(* IEC 61131-3 sources: Palletizer_Control_with_Automation_Studio/Task_1/Logical/Libraries/MpCom, 3 files *)

(* ---- MpCom.typ ---- *)
TYPE
	MpComConfigScopeEnum :
		(
		mpCOM_CONFIG_SCOPE_COMPONENT := 0, (*Import / Export configuration only for given component*)
		mpCOM_CONFIG_SCOPE_BRANCH := 1 (*Import / Export configuration for given component and all its sub-components*)
		);
	MpComStatusIDType : 	STRUCT
		ID : MpComErrorEnum; (*Status ID*)
		Severity : MpComSeveritiesEnum; (*Status severity*)
		Facility : MpComFacilitiesEnum; (*Status facility*)
		Code : UINT; (*Status / Error code*)
	END_STRUCT;
	MpComDiagType : 	STRUCT
		StatusID : MpComStatusIDType; (*StatusID diagnostic structure *)
	END_STRUCT;
	MpComConfigManagerInfoType : 	STRUCT
		Diag : MpComDiagType; (*Diagnostic structure for the status ID*)
	END_STRUCT;
	MpComDumpInternalType : 	STRUCT
		CmdOld : BOOL;
	END_STRUCT;
	MpComLoggerUISetupType : 	STRUCT
		LoggerListSize : UINT := 20; (*Number of logger entries to be displayed on one page of the list in the HMI application*)
		LoggerScrollWindow : USINT := 0; (*Determines how many entries from the list are displayed in advance when scrolling up and down*)
	END_STRUCT;
	MpComLoggerUIConnectType : 	STRUCT
		Status : MpComLoggerUIStatusEnum;
		List : MpComLoggerUILoggerListType; (*List of resultant logger entries*)
		Clear : BOOL; (*Clean the internal buffer*)
		SearchFilter : STRING[255]; (*Filter used to define the visibility of entries*)
	END_STRUCT;
	MpComLoggerUIStatusEnum :
		(
		mpCOM_LOGGERUI_IDLE := 0,
		mpCOM_LOGGERUI_REFRESH := 1,
		mpCOM_LOGGERUI_ERROR := 2
		);
	MpComLoggerUILoggerListType : 	STRUCT
		Message : ARRAY[0..19]OF STRING[255]; (*List of logger entries: message*)
		StatusID : ARRAY[0..19]OF DINT; (*List of logger entries: status ID*)
		ErrorNumber : ARRAY[0..19]OF UINT; (*List of logger entries: error code as part of Status ID*)
		Time : ARRAY[0..19]OF MpComLoggerUIDateTimeType; (*List of logger entries: date, time and microseconds*)
		Component : ARRAY[0..19]OF STRING[50]; (*List of logger entries: component name*)
		Facility : ARRAY[0..19]OF MpComFacilitiesEnum; (*List of logger entries: facility as part of Status ID*)
		Severity : ARRAY[0..19]OF MpComSeveritiesEnum; (*List of logger entries: severity as part of Status ID*)
		PageUp : BOOL; (*Jumps to the start of the current page and then scrolls up one page at a time *)
		PageDown : BOOL; (*Jumps to the end of the current page and then scrolls down one page at a time *)
		StepUp : BOOL; (*Selects the previous entry in the list*)
		StepDown : BOOL; (*Selects the next entry in the list*)
		RangeStart : REAL; (*Shows a bar indicating which part of the list is currently being displayed-Start [%]*)
		RangeEnd : REAL; (*Shows a bar indicating which part of the list is currently being displayed-End [%]*)
	END_STRUCT;
	MpComLoggerUIDateTimeType : 	STRUCT
		DateTime : DATE_AND_TIME; (*List of logger entries: date and time: the view could be customized on VC*)
		Microseconds : UDINT; (*List of logger entries: additional information about microseconds when the event was triggered*)
	END_STRUCT;
	MpComLoggerUIInfoType : 	STRUCT
		CurrentBufferEntries : UINT; (*Number of entries currently in the internal buffer. It is a ring buffer, it means that reached the BufferSize it doesn't increase any more*)
		Diag : MpComDiagType; (*Diagnostic structure for the status ID*)
	END_STRUCT;
END_TYPE

(* ---- MpComError.typ ---- *)
TYPE
    MpComErrorEnum :
        ( (* Error numbers of library MpCom *)
        mpCOM_NO_ERROR := 0, (* No error *)
        mpCOM_ERR_ACTIVATION := -1064239103, (* Could not create component [Error: 1, 0xc0910001] *)
        mpCOM_ERR_MPLINK_NULL := -1064239102, (* MpLink is NULL pointer [Error: 2, 0xc0910002] *)
        mpCOM_ERR_MPLINK_INVALID := -1064239101, (* MpLink connection not allowed [Error: 3, 0xc0910003] *)
        mpCOM_ERR_MPLINK_CHANGED := -1064239100, (* MpLink modified [Error: 4, 0xc0910004] *)
        mpCOM_ERR_MPLINK_CORRUPT := -1064239099, (* Invalid MpLink contents [Error: 5, 0xc0910005] *)
        mpCOM_ERR_LINK_NOT_POSSIBLE := -1064238848, (* Connection not possible [Error: 256, 0xc0910100] *)
        mpCOM_ERR_FILE_SYSTEM := -1064238847, (* Error editing file [Error: 257, 0xc0910101] *)
        mpCOM_ERR_INVALID_FILE_DEV := -1064238846, (* Invalid file device [Error: 258, 0xc0910102] *)
        mpCOM_ERR_INVALID_FILE_NAME := -1064238845, (* Invalid filename [Error: 259, 0xc0910103] *)
        mpCOM_ERR_NO_CONFIG_IMPORT := -1064238844, (* No configuration data was imported [Error: 260, 0xc0910104] *)
        mpCOM_ERR_MISSING_UICONNECT := -1064238843, (* Missing value on UIConnect [Error: 261, 0xc0910105] *)
        mpCOM_ERR_CONFIG_IMPORT_ERR := -1064238842, (* A syntax error was detected in the config-import file [Error: 262, 0xc0910106] *)
        mpCOM_ERR_WRONG_FILTER_STRING := -1064238841, (* Error in the filter string [Error: 263, 0xc0910107] *)
        mpCOM_ERR_COMPONENT_NOT_FOUND := -1064238840 (* The given mapp-component was not found [Error: 264, 0xc0910108] *)
        );
END_TYPE

(* ---- MpCom.fun ---- *)
FUNCTION_BLOCK MpComConfigManager (*Export / Import configuration data*) (* $GROUP=mapp Services,$CAT=mapp Link,$GROUPICON=Icon_mapp.png,$CATICON=Icon_MpCom.png *)
	VAR_INPUT
		MpLink : REFERENCE TO MpComIdentType; (*Incoming communication handle (map standard interface)*) (* *) (*#PAR#;*)
		Enable : BOOL; (*Enables/Disables the function block (mapp standard interface)*) (* *) (*#PAR#;*)
		ErrorReset : BOOL; (*Resets all function block errors (mapp standard interface)*) (* *) (*#PAR#;*)
		DeviceName : REFERENCE TO STRING[50]; (*Name of device where file should be created*) (* *) (*#CMD#;*)
		FileName : REFERENCE TO STRING[255]; (*Name of file to import / create*) (* *) (*#CMD#;*)
		Scope : MpComConfigScopeEnum; (*Scope of configuration to export/import*) (* *) (*#CMD#;*)
		Export : BOOL; (*Export configuration to XML-File*) (* *) (*#CMD#;*)
		Import : BOOL; (*Import configuration from XML-File*) (* *) (*#CMD#;*)
	END_VAR
	VAR_OUTPUT
		Active : BOOL; (*Function block is active (mapp standard interface)*) (* *) (*#PAR#;*)
		Error : BOOL; (*Indicates an error (mapp standard interface)*) (* *) (*#PAR#;*)
		StatusID : DINT; (*Error/Status information (mapp standard interface)*) (* *) (*#PAR#;*)
		CommandBusy : BOOL; (*Function block is busy processing a command*) (* *) (*#CMD#OPT#;*)
		CommandDone : BOOL; (*Command is finished*) (* *) (*#CMD#;*)
		Info : MpComConfigManagerInfoType; (*Additional information about the component*) (* *) (*#CMD#;*)
	END_VAR
	VAR
		Internal : {REDUND_UNREPLICABLE} MpComConfigInternalType; (*Internal data*)
	END_VAR
END_FUNCTION_BLOCK

FUNCTION_BLOCK MpComLoggerUI (*Get mapp logger information*) (* $GROUP=mapp Services,$CAT=mapp Link,$GROUPICON=Icon_mapp.png,$CATICON=Icon_MpCom.png *)
	VAR_INPUT
		MpLink : REFERENCE TO MpComIdentType; (*Incoming communication handle (map standard interface)*) (* *) (*#PAR#;*)
		Enable : BOOL; (*Enables/Disables the function block (mapp standard interface)*) (* *) (*#PAR#;*)
		ErrorReset : BOOL; (*Resets all function block errors (mapp standard interface)*) (* *) (*#PAR#;*)
		Scope : MpComConfigScopeEnum; (*Scope of configuration to export/import*) (* *) (*#PAR#;*)
		EntryFilter : STRING[255]; (*Scope filter to define which entries will be part of the internal logger*) (* *) (*#PAR#;OPT#;*)
		BufferSize : UINT; (*Size of the internal buffer (0=default size 100)*) (* *) (*#PAR#;OPT#;*)
		UISetup : MpComLoggerUISetupType; (*Used to configure the elements connected to the HMI application*) (* *) (*#PAR#;*)
		UIConnect : REFERENCE TO MpComLoggerUIConnectType; (*This structure contains the parameters needed for the connection to the HMI application*) (* *) (*#CMD#;*)
		Clear : BOOL; (*Delete all entries inside the internal buffer*) (* *) (*#CMD#;OPT#;*)
	END_VAR
	VAR_OUTPUT
		Active : BOOL; (*Function block is active (mapp standard interface)*) (* *) (*#PAR#;*)
		Error : BOOL; (*Indicates an error (mapp standard interface)*) (* *) (*#PAR#;*)
		StatusID : DINT; (*Error/Status information (mapp standard interface)*) (* *) (*#PAR#; *)
		Info : MpComLoggerUIInfoType; (*Additional information about the component*) (* *) (*#CMD#;*)
	END_VAR
	VAR
		Internal : {REDUND_UNREPLICABLE} MpComInternalDataType; (*Internal data*) (* *) (*#OMIT#;*)
	END_VAR
END_FUNCTION_BLOCK

FUNCTION MpComLink : DINT (*Creates a hierarchy for the mapp components*) (* $GROUP=mapp Services,$CAT=mapp Link,$GROUPICON=Icon_mapp.png,$CATICON=Icon_MpCom.png *)
	VAR_INPUT
		ParentLink : MpComIdentType; (*Link to parent*) (* *) (*#PAR#;*)
		MpLink : MpComIdentType; (*Link to mapp-component*) (* *) (*#PAR#;*)
	END_VAR
END_FUNCTION

FUNCTION_BLOCK MpComLinkToParent (*Creates a hierarchy for the mapp components*) (* $GROUP=mapp Services,$CAT=mapp Link,$GROUPICON=Icon_mapp.png,$CATICON=Icon_MpCom.png *)
	VAR_INPUT
		ParentLink : MpComIdentType; (*Link to parent*) (* *) (*#PAR#;*)
		MpLink : REFERENCE TO MpComIdentType; (*Link to mapp-component*) (* *) (*#PAR#;*)
	END_VAR
	VAR_OUTPUT
		LinkOut : {REDUND_UNREPLICABLE} MpComIdentType; (*Outgoing component link (MpLink)*) (* *) (*#PAR#;*)
		StatusID : DINT; (*Error output*) (* *) (*#PAR#;*)
	END_VAR
END_FUNCTION_BLOCK

FUNCTION_BLOCK MpComDump (*Creates a mapp diagnostic dump file*) (* $GROUP=mapp Services,$CAT=mapp Link,$GROUPICON=Icon_mapp.png,$CATICON=Icon_MpCom.png *)
	VAR_INPUT
		Enable : BOOL; (*Enables/Disables the function block *) (* *) (*#PAR#;*)
		Dump : BOOL; (*A positive signal on this input triggers a dump*) (* *) (*#CMD#;*)
		DeviceName : STRING[20]; (*Name of device where file should be created*) (* *) (*#CMD#;*)
		FileName : STRING[40]; (*Name of file to create*) (* *) (*#CMD#;*)
	END_VAR
	VAR_OUTPUT
		Active : BOOL; (*Function block is active (enabled)*) (* *) (*#PAR#;*)
		Error : BOOL; (*A error has occurred during the last operation*) (* *) (*#PAR#;*)
		StatusID : DINT; (*Information about the error that has occurred*) (* *) (*#PAR#;*)
		CommandBusy : BOOL; (*Function block is busy processing a command*) (* *) (*#CMD#OPT#;*)
		CommandDone : BOOL; (*Command is finished*) (* *) (*#CMD#;*)
	END_VAR
	VAR
		Internal : {REDUND_UNREPLICABLE} MpComDumpInternalType;
	END_VAR
END_FUNCTION_BLOCK

FUNCTION_BLOCK MpComGetLink (*Get MpLink by component name*)
	VAR_INPUT
		Enable : BOOL; (*Enables/Disables the function block *) (* *) (*#PAR#;*)
		ComponentName : REFERENCE TO STRING[100]; (*Full-qualified component name (including scope if necessary)*) (* *) (*#CMD#;*)
	END_VAR
	VAR_OUTPUT
		MpLink : {REDUND_UNREPLICABLE} MpComIdentType; (*Link to mapp-component*) (* *) (*#CMD#;*)
		Error : BOOL; (*A error has occurred when trying to find component*) (* *) (*#PAR#;*)
		Active : BOOL; (*Component was found (MpLink valid)*) (* *) (*#PAR#;*)
		StatusID : DINT; (*Information about the error that has occurred*) (* *) (*#PAR#;*)
	END_VAR
	VAR
		Internal : {REDUND_UNREPLICABLE} BOOL;
	END_VAR
END_FUNCTION_BLOCK
